Fanuc KAREL source: KO00021.KL

PROGRAM KO00021
%NOLOCKGROUP
VAR
  P1: XYZWPREXT
  P2: XYZWPREXT
  P3: XYZWPREXT
  P4: XYZWPREXT
  OUT: POSITION
BEGIN
  OUT = FRAME(P1, P2, P3, P4)
END KO00021
